// TIA Portal V20 export
FUNCTION_BLOCK "05_Not-Aus"   // FB44, FBD
TITLE = NOT-HALT Funktionen
{ S7_Optimized_Access := 'TRUE' }
// stored: MemoryReserve 100, SetENOAutomatically false
BEGIN

NETWORK
TITLE = NOT-HALT Baustein bearbeiten?
      AN    "03_Betriebsart_DB"."NOT-HALT OK";
      JCN   ENDE;


NETWORK
TITLE = Setzen Signal Richten erforderlich nach NOT-HALT

NETWORK
TITLE = Rücksetzen der Freigaben aus Automatik/Manuell/Einfädeln

NETWORK
TITLE = E-Freigaben Rücksetzen

NETWORK
TITLE = Rücksetzen der Ausgänge

NETWORK
TITLE = Rücksetzen der Zeiten

NETWORK
TITLE = Rücksetzen aller Antriebsfreigaben
// Freigaben werden im Antriebsbaustein entzogen







NETWORK
TITLE = Übergabe Position in NOT-HALT um Lage stabil zu halten

NETWORK
TITLE = Setzen von Systeminitialiesierung

NETWORK
TITLE = Rücksetzen der Betriebsarten
//      SET
//      R     "HMI_Signale".Ablauf_aktiv
//      R     "HMI_Signale".Automatik_BA
//      R     "HMI_Signale".Manuell_BA
//      R     "HMI_Signale".Verwalten_BA
//      R     "HMI_Signale".Richten_BA
//      R     "HMI_Signale".Stop_nach_Zyklus

NETWORK
TITLE = Betriebsart Einzelbetrieb
//      SET
//      R     "HMI_Signale".Dauer_Manuell_Betrieb

NETWORK
TITLE = Rücksetze Störmeldungen im NOT-HALT
//      L     0
//      T     DB512.DBD    4
//      T     DB512.DBD    8
//      T     DB512.DBD   12
//      T     DB512.DBD   16


NETWORK
TITLE = 
ENDE: NOP   0;

END_FUNCTION_BLOCK
